(* IEC 61131-3 sources: ae-safety-with-tia-fplc/src, 5 files *)

(* ---- ConveyorTypes.st ---- *)
NAMESPACE SimpleConveyor

    TYPE conveyorInputs:
        STRUCT
            SafetyOK          : BOOL; // Single safety signal from safety relay line
            StartButton       : BOOL; // Manual start button
            StopButton        : BOOL; // Manual stop button
            ItemAtPosA        : BOOL; // Sensor: Item at Position A
            ItemAtPosB        : BOOL; // Sensor: Item at Position B
            ConveyorRunning   : BOOL; // Feedback: Motor running
            MotorFault        : BOOL; // Motor fault signal
            MaxCounterValue   : INT := 10; // Maximum counter value
        END_STRUCT;
    END_TYPE

    TYPE conveyorOutputs:
        STRUCT
            ConveyorMotor     : BOOL; // Conveyor motor control
            StatusLED_Green   : BOOL; // System OK indicator
            StatusLED_Red     : BOOL; // System fault indicator
            StatusLED_Yellow  : BOOL; // System warning/starting
            AlarmHorn         : BOOL; // Safety alarm
            SystemState       : INT; // Current system state
            ItemCounter       : INT; // Current item counter
            FaultCode         : INT; // Active fault code
        END_STRUCT;
    END_TYPE

END_NAMESPACE

(* ---- tcpCommunication.st ---- *)
USING Siemens.Simatic.Communication.Ouc;

TYPE connectionResult:
    STRUCT
        connected : BOOL;
        dataReceived : BOOL;
        receiveStatus : WORD;
        data0 : BYTE;
        data1 : BYTE;
        safetySignal : BOOL;
        connectionError : BOOL;
        connectionStatus : WORD;
    END_STRUCT;
END_TYPE
CLASS SafetySignalReceiver
    VAR PRIVATE
        _connectionConfig : ConnectionConfiguration := (
            ConnectionID := WORD#16#1,
            ActiveEstablished := FALSE,
            LocalPort := UINT#2001,
            ConnectionType := BYTE#16#0B  // TCP
        );
        _connection : Connect;
        _receive : TcpReceive;

        _safetySignal : Bool := FALSE;
        _connected : Bool := FALSE;
        _data : ARRAY[0..1] OF BYTE;  // Buffer for received data

        //Debug variables
        _lastData0 : BYTE;  // For debugging
        _lastData1 : BYTE;  // For debugging
        _receiveStatus : WORD;  // For debugging
        _dataReceived : BOOL;  // For debugging
        _dataEverReceived : BOOL := FALSE; //Track if data has been ever received
    END_VAR

    METHOD PUBLIC Execute : Bool
        // Connection management - runs every cycle like in example
        _connection(
            execute := NOT _connected AND NOT _connection.busy,
            connectionID := _connectionConfig.ConnectionID,
            connectionConfiguration := _connectionConfig
        );

        IF _connection.done THEN
            _connected := TRUE;
        END_IF;

        // Receive data if connected - just like example
        IF _connected THEN
            _receive(
                enable := TRUE,
                connectionID := _connectionConfig.ConnectionID,
                adhocMode := TRUE,  // Use adhoc mode like in the example
                data := _data
            );

            // Debug info
            _receiveStatus := _receive.status;
            _dataReceived := _receive.newDataReceived;

            // Process data when received
            IF _receive.newDataReceived THEN
                _lastData0 := _data[0];
                _lastData1 := _data[1];
                _safetySignal := (_data[0] > BYTE#0);  // Only checking first byte for now
                _dataEverReceived := TRUE; //Set flag when data is received
                _dataReceived := TRUE; //Current Cycle has data
            ELSE
                _dataReceived := FALSE; //Reset for current cycle
            END_IF;
        END_IF;

        Execute := _safetySignal;
    END_METHOD

    METHOD PUBLIC GetDebugInfo : connectionResult
        VAR
            result : connectionResult;
        END_VAR
        result.connected := _connected;
        result.dataReceived := _dataReceived OR _dataEverReceived;
        result.receiveStatus := _receiveStatus;
        result.data0 := _lastData0;
        result.data1 := _lastData1;
        result.safetySignal := _safetySignal;
        result.connectionError := _connection.error;
        result.connectionStatus := _connection.status;

        GetDebugInfo := result;

    END_METHOD
END_CLASS

(* ---- conveyorControl.st ---- *)
USING System.Timer;

NAMESPACE SimpleConveyor

    CLASS ConveyorController
        VAR PUBLIC
            Inputs : conveyorInputs;
            Outputs : conveyorOutputs;
        END_VAR

        VAR PRIVATE
            SystemEnabled       : BOOL := FALSE;
            ConveyorCommand     : BOOL := FALSE;
            ItemCounter         : INT := 0;
            CounterDirection    : BOOL := TRUE;
            CurrentState        : INT := 0; // 0=STOPPED, 1=STARTING, 2=RUNNING, 3=FAULT

            // Edge detection
            ItemAtPosB_Old      : BOOL := FALSE;
            StartButton_Old     : BOOL := FALSE;
            StopButton_Old      : BOOL := FALSE;
            SafetyOK_Old        : BOOL := FALSE;

            // Timers
            StartDelay          : OnDelay;
            SafetyLossTimer     : OnDelay; // Timer to monitor safety signal loss

            // Safety monitoring
            SafetyLossDetected  : BOOL := FALSE;
            SafetyRestored      : BOOL := FALSE;
        END_VAR

        METHOD PUBLIC Execute
            THIS.CheckSafety();
            THIS.ProcessButtons();
            THIS.HandleStateMachine();
            THIS.ProcessItems();
            THIS.SetOutputs();

            // Store previous safety state
            THIS.SafetyOK_Old := THIS.Inputs.SafetyOK;
        END_METHOD

        METHOD PRIVATE CheckSafety
            VAR
                SafetyFalling   : BOOL;
                SafetyRising    : BOOL;
            END_VAR

            // Detect safety signal transitions
            SafetyFalling := NOT THIS.Inputs.SafetyOK AND THIS.SafetyOK_Old;
            SafetyRising := THIS.Inputs.SafetyOK AND NOT THIS.SafetyOK_Old;

            // Monitor safety signal loss
            IF SafetyFalling THEN
                THIS.SafetyLossDetected := TRUE;
                THIS.SafetyLossTimer(signal := TRUE, duration := T#5s); // Start monitoring timer
            END_IF;

            // Check if safety has been restored
            IF SafetyRising THEN
                THIS.SafetyRestored := TRUE;
                THIS.SafetyLossDetected := FALSE;
                THIS.SafetyLossTimer(signal := FALSE);
            END_IF;

            // Basic safety check
            IF THIS.Inputs.SafetyOK  AND NOT THIS.Inputs.MotorFault THEN
                THIS.SystemEnabled := TRUE;
                IF THIS.CurrentState = 3 AND This.SafetyRestored THEN
                    THIS.CurrentState := 0; // Go to stopped when safety restored
                    THIS.SafetyRestored := FALSE; // Reset flag
                END_IF;
            ELSE
                THIS.SystemEnabled := FALSE;
                THIS.CurrentState := 3; // Fault state
            END_IF;

            // Extended safety loss handling
            IF THIS.SafetyLossTimer.output THEN
                THIS.Outputs.FaultCode := 3; // Extended safety loss fault
            END_IF;
        END_METHOD

        METHOD PRIVATE ProcessButtons
            VAR
                StartEdge : BOOL;
                StopEdge : BOOL;
            END_VAR

            // Edge detection for buttons
            StartEdge := THIS.Inputs.StartButton AND NOT THIS.StartButton_Old;
            StopEdge := THIS.Inputs.StopButton AND NOT THIS.StopButton_Old;
            THIS.StartButton_Old := THIS.Inputs.StartButton;
            THIS.StopButton_Old := THIS.Inputs.StopButton;

            // Start logic: Only if safety OK and system stopped
            IF StartEdge AND THIS.SystemEnabled AND THIS.CurrentState = 0 THEN
                THIS.CurrentState := 1; // Start
            END_IF;

            // Stop logic: Always stop if button pressed or safety not OK
            IF StopEdge OR NOT THIS.SystemEnabled THEN
                THIS.CurrentState := 0; // Stop
                THIS.StartDelay(signal := FALSE); // Reset start timer
            END_IF;
        END_METHOD

        METHOD PRIVATE HandleStateMachine
            CASE THIS.CurrentState OF
                0: // STOPPED
                    THIS.ConveyorCommand := FALSE;

                1: // STARTING
                    // Only allow starting if safety is stable
                    IF NOT THIS.SafetyLossDetected THEN
                        THIS.StartDelay(signal := TRUE, duration := T#2S);
                        IF THIS.StartDelay.output THEN
                            THIS.CurrentState := 2; // Running
                            THIS.StartDelay(signal := FALSE);
                        END_IF;
                    ELSE
                        THIS.CurrentState := 0; // Return to stopped if safety unstable
                    END_IF;
                2: // RUNNING
                    THIS.ConveyorCommand := TRUE;

                3: // FAULT
                    THIS.ConveyorCommand := FALSE;
                    // Can only exit fault by fixing safety and pressing start
                    // Additional safety recovery logic
                    IF THIS.SafetyRestored AND THIS.Inputs.SafetyOK THEN
                        // Wait for explicit restart after safety restoration
                        THIS.Outputs.StatusLED_Yellow := TRUE; // Indicate ready for restart
                    END_IF;
            END_CASE;
        END_METHOD

        METHOD PRIVATE ProcessItems
            VAR
                ItemEdge : BOOL;
            END_VAR

            // Edge detection for item at Position B
            ItemEdge := THIS.Inputs.ItemAtPosB AND NOT THIS.ItemAtPosB_Old;
            THIS.ItemAtPosB_Old := THIS.Inputs.ItemAtPosB;

            // Counter logic - only when RUNNING and item detected
            IF THIS.CurrentState = 2 AND ItemEdge THEN // Running and item detected
                IF THIS.CounterDirection THEN
                    // Counting UP
                    THIS.ItemCounter := THIS.ItemCounter + 1;
                    IF THIS.ItemCounter >= THIS.Inputs.MaxCounterValue THEN
                        THIS.CounterDirection := FALSE; //Switch to count down
                    END_IF;
                ELSE
                    THIS.ItemCounter := THIS.ItemCounter - 1;
                    IF THIS.ItemCounter <= 0 THEN
                        THIS.CounterDirection := TRUE; //Swithc to count up
                    END_IF;
                END_IF;
            END_IF;
        END_METHOD

        METHOD PRIVATE SetOutputs
            // Motor control with safety
            THIS.Outputs.ConveyorMotor := THIS.ConveyorCommand AND THIS.SystemEnabled;

            // Status LEDs with enhanced safety indication
            THIS.Outputs.StatusLED_Green := (THIS.CurrentState = 2);  // Running = Green
            THIS.Outputs.StatusLED_Red := (THIS.CurrentState = 3) OR THIS.SafetyLossDetected;    // Fault = Red
            THIS.Outputs.StatusLED_Yellow := (THIS.CurrentState = 1) OR (THIS.SafetyRestored AND THIS.CurrentState = 3); // Starting or Ready for Restart = Yellow

            // Alarm
            THIS.Outputs.AlarmHorn := (THIS.CurrentState = 3) OR (THIS.SafetyLossDetected AND THIS.SafetyLossTimer.output);

            // Status info
            THIS.Outputs.SystemState := THIS.CurrentState;
            THIS.Outputs.ItemCounter := THIS.ItemCounter;

            // Fault code assignment
            IF THIS.CurrentState = 3 THEN
                IF THIS.SafetyLossDetected AND THIS.SafetyLossTimer.output THEN
                    THIS.Outputs.FaultCode := 3; // Extended safety loss
                ELSIF NOT THIS.Inputs.SafetyOK THEN
                    THIS.Outputs.FaultCode := 1; // Safety fault
                ELSIF THIS.Inputs.MotorFault THEN
                    THIS.Outputs.FaultCode := 2; // Motor fault
                ELSE
                    THIS.Outputs.FaultCode := 1; // General safety fault
                END_IF;
            ELSE
                THIS.Outputs.FaultCode := 0; // No fault
            END_IF;
        END_METHOD

    END_CLASS
END_NAMESPACE

(* ---- configuration.st ---- *)
USING SimpleConveyor;
CONFIGURATION MyConfiguration
    TASK Main(Priority := 1);

    PROGRAM P1 WITH Main: ConveyorControl;

    VAR_GLOBAL
        // Physical Input I/O

        // Moved from defined Input Card for Simulation
        // IO_StartButton       AT %IX0.1 : BOOL;
        // IO_StopButton        AT %IX0.2 : BOOL;
        // IO_ItemAtPosA        AT %IX0.3 : BOOL;
        // IO_ItemAtPosB        AT %IX0.4 : BOOL;
        // IO_ConveyorRunning   AT %IX0.5 : BOOL;
        // IO_MotorFault        AT %IX0.6 : BOOL;

        IO_StartButton       AT %IX4.1 : BOOL;
        IO_StopButton        AT %IX4.2 : BOOL;
        IO_ItemAtPosA        AT %IX4.3 : BOOL;
        IO_ItemAtPosB        AT %IX4.4 : BOOL;
        IO_ConveyorRunning   AT %IX4.5 : BOOL;
        IO_MotorFault        AT %IX4.6 : BOOL;
        IO_MaxCounterValue   AT %IW2 : INT;

        // Physical Output I/O
        // Moved from defined Output Card for Simulation

        // IO_ConveyorMotor     AT %QX0.0 : BOOL;
        // IO_StatusLED_Green   AT %QX0.2 : BOOL;
        // IO_StatusLED_Red     AT %QX0.3 : BOOL;
        // IO_StatusLED_Yellow  AT %QX0.4 : BOOL;
        // IO_AlarmHorn         AT %QX0.5 : BOOL;

        IO_ConveyorMotor     AT %QX8.0 : BOOL;
        IO_StatusLED_Green   AT %QX8.2 : BOOL;
        IO_StatusLED_Red     AT %QX8.3 : BOOL;
        IO_StatusLED_Yellow  AT %QX8.4 : BOOL;
        IO_AlarmHorn         AT %QX8.5 : BOOL;
        IO_SystemState       AT %QW2 : INT;
        IO_ItemCounter       AT %QW4 : INT;
        IO_FaultCode         AT %QW6 : INT;

        // Conveyor instance
        Conveyor : ConveyorController;

        //Safety communication instance
        SafetyComm : SafetySignalReceiver;

        //debug Instance

        debugInfo : connectionResult;
END_VAR
END_CONFIGURATION

(* ---- MainProgram.st ---- *)
USING SimpleConveyor;
USING Siemens.Simatic.Communication.OUC;

PROGRAM ConveyorControl
    VAR_EXTERNAL
         // Reference to global input I/O variables
         //IO_SafetyOK          : BOOL;
         IO_StartButton       : BOOL;
         IO_StopButton        : BOOL;
         IO_ItemAtPosA        : BOOL;
         IO_ItemAtPosB        : BOOL;
         IO_ConveyorRunning   : BOOL;
         IO_MotorFault        : BOOL;
         IO_MaxCounterValue   : INT;

         // Reference to global output I/O variables
         IO_ConveyorMotor     : BOOL;
         IO_StatusLED_Green   : BOOL;
         IO_StatusLED_Red     : BOOL;
         IO_StatusLED_Yellow  : BOOL;
         IO_AlarmHorn         : BOOL;
         IO_SystemState       : INT;
         IO_ItemCounter       : INT;
         IO_FaultCode         : INT;

         //Classes instances reference of the global
         Conveyor : ConveyorController;
         SafetyComm : SafetySignalReceiver;
         debugInfo : connectionResult;
    END_VAR
    VAR
        FirstCycle : BOOL := TRUE;
    END_VAR

    // // Initialize TCP communications on first cycle
    // IF FirstCycle THEN
    //     SafetyComm.Configure();
    //     FirstCycle := FALSE;
    // END_IF;

    //Get debug info
    debugInfo := SafetyComm.GetDebugInfo();
    // Map inputs
    //Conveyor.Inputs.SafetyOK := IO_SafetyOK;
    Conveyor.Inputs.SafetyOK := SafetyComm.Execute(); // Get safety signal via TCP
    Conveyor.Inputs.StartButton := IO_StartButton;
    Conveyor.Inputs.StopButton := IO_StopButton;
    Conveyor.Inputs.ItemAtPosA := IO_ItemAtPosA;
    Conveyor.Inputs.ItemAtPosB := IO_ItemAtPosB;
    Conveyor.Inputs.ConveyorRunning := IO_ConveyorRunning;
    Conveyor.Inputs.MotorFault := IO_MotorFault;
    Conveyor.Inputs.MaxCounterValue := IO_MaxCounterValue;

    // Execute conveyor logic
    Conveyor.Execute();

    // Map outputs
    IO_ConveyorMotor := Conveyor.Outputs.ConveyorMotor;
    IO_StatusLED_Green := Conveyor.Outputs.StatusLED_Green;
    IO_StatusLED_Red := Conveyor.Outputs.StatusLED_Red;
    IO_StatusLED_Yellow := Conveyor.Outputs.StatusLED_Yellow;
    IO_AlarmHorn := Conveyor.Outputs.AlarmHorn;
    IO_SystemState := Conveyor.Outputs.SystemState;
    IO_ItemCounter := Conveyor.Outputs.ItemCounter;
    IO_FaultCode := Conveyor.Outputs.FaultCode;

END_PROGRAM
